(* IEC 61131-3 sources: FACTORY_io/fabrica-viva/etapa-3, 3 files *)

(* ---- fragmento-bloques.st ---- *)
(* ===== Etapa 3 · Bloque de función FB_Cola =====
   Una cola FIFO de códigos: lo primero que entra es lo primero que sale. Complétalo con un ARRAY.
   - Meter (un pulso): añade Valor al final de la cola.
   - Sacar (un pulso): quita el primero de la cola.
   - Si llegan los dos en el mismo ciclo, primero se saca y después se mete.
   - Primero: el valor que está a la cabeza (0 si la cola está vacía). Cantidad: cuántos hay. *)
FUNCTION_BLOCK FB_Cola
VAR_INPUT
  Meter : BOOL;
  Valor : DINT;
  Sacar : BOOL;
END_VAR
VAR_OUTPUT
  Primero : DINT;
  Cantidad : INT;
END_VAR
VAR
  Datos : ARRAY[0..15] OF DINT;   (* hasta 16 cajas en cola *)
  (* tus variables internas del bloque *)
END_VAR

(* ---- tu código del bloque ---- *)
END_FUNCTION_BLOCK

(* ---- solucion.st ---- *)
(* Fábrica viva · Etapa 3 · Solución de referencia: colas FIFO con ARRAY para clasificar por código. *)
FUNCTION_BLOCK FB_Cola
VAR_INPUT
  Meter : BOOL;
  Valor : DINT;
  Sacar : BOOL;
END_VAR
VAR_OUTPUT
  Primero : DINT;
  Cantidad : INT;
END_VAR
VAR
  Datos : ARRAY[0..15] OF DINT;
  i : INT;
END_VAR

(* Sacar desplaza todo un puesto hacia la cabeza; meter escribe detrás del último. *)
IF Sacar AND Cantidad > 0 THEN
  FOR i := 0 TO 14 DO
    Datos[i] := Datos[i + 1];
  END_FOR;
  Cantidad := Cantidad - 1;
END_IF;
IF Meter AND Cantidad < 16 THEN
  Datos[Cantidad] := Valor;
  Cantidad := Cantidad + 1;
END_IF;
IF Cantidad > 0 THEN
  Primero := Datos[0];
ELSE
  Primero := 0;
END_IF;
END_FUNCTION_BLOCK

FUNCTION_BLOCK FB_Cinta
VAR_INPUT
  Habilitar : BOOL;
  Presencia : BOOL;
  Rearme : BOOL;
END_VAR
VAR_OUTPUT
  Motor : BOOL;
  Atasco : BOOL;
END_VAR
VAR
  Tapada : TON;
END_VAR

Tapada(IN := Presencia AND Motor, PT := T#3s);
IF Rearme THEN
  Atasco := FALSE;
END_IF;
IF Tapada.Q THEN
  Atasco := TRUE;
END_IF;
Motor := Habilitar AND NOT Atasco;
END_FUNCTION_BLOCK

VAR_INPUT
  Marcha : BOOL;
  Paro : BOOL;
  Seta : BOOL;
  FotocelulaRecepcion : BOOL;
  CajasRecibidas : INT;
END_VAR
VAR_OUTPUT
  CintaRecepcion : BOOL;
  Alimentador : BOOL;
  Baliza : INT;
END_VAR
VAR
  EnMarcha : BOOL;
END_VAR

VAR_INPUT
  Rearme : BOOL;
  FotocelulaAtasco : BOOL;
  LecturaOk : BOOL;
  CodigoCaja : DINT;
  FotocelulaRechazo : BOOL;
  CajasRechazadas : INT;
  CajasFinLinea : INT;
END_VAR
VAR_OUTPUT
  CintaControl : BOOL;
  Desvio : BOOL;
  AlarmaAtasco : BOOL;
END_VAR
VAR
  Control : FB_Cinta;
  Leida : R_TRIG;
  Llega : R_TRIG;
  SinEtiqueta : BOOL;
  Pendiente : BOOL;
  Retardo : TON;
  Empuje : TP;
END_VAR

VAR_INPUT
  FotocelulaExpres : BOOL;
  FotocelulaDevol : BOOL;
  CajasExpres : INT;
  CajasDevueltas : INT;
  CajasPedidos : INT;
END_VAR
VAR_OUTPUT
  CintaClasificacion : BOOL;
  DesvioExpres : BOOL;
  DesvioDevol : BOOL;
END_VAR
VAR
  ColaA : FB_Cola;
  ColaB : FB_Cola;
  CodigoEnA : DINT;
  LlegaA : R_TRIG;
  LlegaB : R_TRIG;
  PendienteA : BOOL;
  PendienteB : BOOL;
  RetardoA : TON;
  RetardoB : TON;
  EmpujeA : TP;
  EmpujeB : TP;
END_VAR

(* Etapas 1 y 2 *)
EnMarcha := (Marcha OR EnMarcha) AND NOT Paro AND Seta AND NOT AlarmaAtasco;
CintaRecepcion := EnMarcha;
Alimentador := EnMarcha;
Control(Habilitar := EnMarcha, Presencia := FotocelulaAtasco, Rearme := Rearme);
CintaControl := Control.Motor;
AlarmaAtasco := Control.Atasco;
IF NOT Seta THEN
  Baliza := 4;
ELSIF AlarmaAtasco THEN
  Baliza := 6;
ELSIF EnMarcha THEN
  Baliza := 1;
ELSE
  Baliza := 2;
END_IF;
Leida(CLK := LecturaOk);
IF Leida.Q THEN
  SinEtiqueta := CodigoCaja = 0;
END_IF;
Llega(CLK := FotocelulaRechazo);
IF Llega.Q AND SinEtiqueta AND EnMarcha THEN
  Pendiente := TRUE;
END_IF;
Retardo(IN := Pendiente, PT := T#450ms);
IF Retardo.Q OR NOT EnMarcha THEN
  Pendiente := FALSE;
END_IF;
Empuje(IN := Retardo.Q, PT := T#600ms);
Desvio := Empuje.Q AND EnMarcha;

(* Etapa 3. Primero se detectan las llegadas; después se decide con la cabeza de cada cola (el código de la
   caja que acaba de llegar) y por último se actualizan las colas, cada una con una sola llamada por ciclo. *)
CintaClasificacion := EnMarcha;
LlegaB(CLK := FotocelulaDevol);
LlegaA(CLK := FotocelulaExpres);
IF LlegaB.Q AND ColaB.Primero = 104 THEN
  PendienteB := TRUE;
END_IF;
CodigoEnA := ColaA.Primero;
IF LlegaA.Q AND CodigoEnA = 103 THEN
  PendienteA := TRUE;
END_IF;
(* la caja que pasa el empujador exprés sin desviarse entra en la cola del tramo siguiente *)
ColaB(Meter := LlegaA.Q AND ColaA.Cantidad > 0 AND CodigoEnA <> 103, Valor := CodigoEnA, Sacar := LlegaB.Q);
ColaA(Meter := Leida.Q AND CodigoCaja <> 0, Valor := CodigoCaja, Sacar := LlegaA.Q);

RetardoA(IN := PendienteA, PT := T#450ms);
IF RetardoA.Q OR NOT EnMarcha THEN
  PendienteA := FALSE;
END_IF;
EmpujeA(IN := RetardoA.Q, PT := T#600ms);
DesvioExpres := EmpujeA.Q AND EnMarcha;
RetardoB(IN := PendienteB, PT := T#450ms);
IF RetardoB.Q OR NOT EnMarcha THEN
  PendienteB := FALSE;
END_IF;
EmpujeB(IN := RetardoB.Q, PT := T#600ms);
DesvioDevol := EmpujeB.Q AND EnMarcha;

(* ---- fragmento-declaraciones.st ---- *)
(* ===== Etapa 3 · Clasificación: señales nuevas ===== *)
VAR_INPUT
  FotocelulaExpres : BOOL;    (* fotocélula antes del empujador exprés (código 103) *)
  FotocelulaDevol : BOOL;     (* fotocélula antes del empujador de devoluciones (código 104) *)
  CajasExpres : INT;          (* cajas retiradas en la cinta de exprés *)
  CajasDevueltas : INT;       (* cajas retiradas en la cinta de devoluciones *)
  CajasPedidos : INT;         (* cajas de pedido normal (101, 102) al final de la clasificación *)
END_VAR
VAR_OUTPUT
  CintaClasificacion : BOOL;  (* la cinta de clasificación y sus dos laterales *)
  DesvioExpres : BOOL;
  DesvioDevol : BOOL;
END_VAR
VAR
  ColaA : FB_Cola;            (* las cajas entre el lector y el empujador exprés *)
  ColaB : FB_Cola;            (* las cajas entre el empujador exprés y el de devoluciones *)
END_VAR
